// TIA Portal project "python_communication" (V18)

(* hardware
DEVICE "S7-1200 station_1"  S7-1200 Station
   slot 0: "Rack_0"  S7-1200 Rack  Rack  V1.0
   slot 1: "PLC_1"  CPU 1214C DC/DC/Rly  6ES7 214-1HG40-0XB0  V4.6
*)

// ===== PLC "PLC_1"  CPU 1214C DC/DC/Rly =====

VAR_GLOBAL   // PLC tag table "Default tag table"
   "Main_Conveyor_Motor" AT %Q10.0 : Bool;
   "Start_But" AT %I10.0 : Bool;
   "Stop_But" AT %I10.1 : Bool;
   "Start_Mem" AT %M1.0 : Bool;
   "First_Detected_Sensor" AT %I10.2 : Bool;
   "Stop_Mem" AT %M2.0 : Bool;
   "Second_Band_Exit_Sensor" AT %I10.3 : Bool;
   "Second_Band_First_Sensor" AT %I10.4 : Bool;
   "Machine_Sensor" AT %I10.5 : Bool;
   "Move_Z_Mem" AT %M3.0 : Bool;
   "Move_Z" AT %Q10.1 : Bool;
   "Grab_İtem" AT %Q10.2 : Bool;
   "Grab_Mem" AT %M4.0 : Bool;
   "Move_X_Mem" AT %M5.0 : Bool;
   "Move_X" AT %Q10.3 : Bool;
   "Moving_X" AT %I10.6 : Bool;
   "Moving_Z" AT %I10.7 : Bool;
   "Second_Band_Motor" AT %Q10.4 : Bool;
   "Second_Band_Motor_Mem" AT %M6.0 : Bool;
   "Defect_Process_Active" AT %M7.0 : Bool;
   "Corner_Band_Motor" AT %Q10.5 : Bool;
   "Main_Band2_Motor" AT %Q10.6 : Bool;
   "Stack_Light(RED)" AT %Q10.7 : Bool;
   "Stack_Light(GREEN)" AT %Q11.0 : Bool;
   "Stack_Light(YELLOW)" AT %Q11.1 : Bool;
   "Python_Alive" AT %M8.0 : Bool;
END_VAR

DATA_BLOCK "DB_Python"   // DB1
{ S7_Optimized_Access := 'FALSE' }
VERSION : 0.1
   VAR
      Trigger : Bool;
      Part_At_Camera : Bool;
      Heartbeat : Bool;
      DefectCount : Int;
      ConfidenceScore : Real;
   END_VAR
BEGIN
END_DATA_BLOCK

// folder: System blocks/Program resources

DATA_BLOCK "timer5"   // DB2
{ S7_Optimized_Access := 'TRUE' }
AUTHOR : Simatic
FAMILY : IEC
NAME : IEC_TMR
VERSION : 1.0
// stored: InstanceOfName IEC_TIMER
"IEC_TIMER"
BEGIN
END_DATA_BLOCK

DATA_BLOCK "timer1"   // DB3
{ S7_Optimized_Access := 'TRUE' }
AUTHOR : Simatic
FAMILY : IEC
NAME : IEC_TMR
VERSION : 1.0
// stored: InstanceOfName IEC_TIMER
"IEC_TIMER"
BEGIN
END_DATA_BLOCK

DATA_BLOCK "Timer2"   // DB4
{ S7_Optimized_Access := 'TRUE' }
AUTHOR : Simatic
FAMILY : IEC
NAME : IEC_TMR
VERSION : 1.0
// stored: InstanceOfName IEC_TIMER
"IEC_TIMER"
BEGIN
END_DATA_BLOCK

DATA_BLOCK "timer3"   // DB5
{ S7_Optimized_Access := 'TRUE' }
AUTHOR : Simatic
FAMILY : IEC
NAME : IEC_TMR
VERSION : 1.0
// stored: InstanceOfName IEC_TIMER
"IEC_TIMER"
BEGIN
END_DATA_BLOCK

// folder: (top level)

FUNCTION "MHJ-PLC-Lab-Function-S71200" : Void   // FC9000, SCL
{ S7_Optimized_Access := 'TRUE' }
VERSION : 0.1
   VAR_TEMP
      rdTimeReturn : Int;
      outputTime : DTL;
      SyncVal : Byte;
      forVal : Int;
      forVal_2 : Int;
      Value : Byte;
   END_VAR
   VAR CONSTANT
      CompVal : Byte := 16#34;
      Value_01 : Byte := 16#11;
      Value_01_DW : DWord := 16#A165_D992;
      Value_02_DW : DWord := 16#58BE_4401;
   END_VAR
BEGIN

   #Value:=PEEK(area := 16#82,
        dbNumber := 0,
        byteOffset := 511);
   #Value := #Value + 1;

   POKE(area := 16#82,
        dbNumber := 0,
        byteOffset := 511,
        value := #Value);

   POKE(area:=16#81,
        dbNumber:=0,
        byteOffset:=1016,
        value:=#Value_01_DW);
   POKE(area := 16#81,
        dbNumber := 0,
        byteOffset := 1020,
        value := #Value_02_DW);

   POKE(area := 16#81,
        dbNumber := 0,
        byteOffset := 511,
        value := B#16#00);

   FOR #forVal := 0 TO 120 DO
       FOR #forVal_2:=0 TO 10 DO
           #rdTimeReturn:=RD_SYS_T(#outputTime);
           #rdTimeReturn := WR_SYS_T(#outputTime);
           #rdTimeReturn := RD_SYS_T(#outputTime);
           #rdTimeReturn := WR_SYS_T(#outputTime);
       END_FOR;
       #SyncVal:= PEEK(area := 16#81,
                      dbNumber := 0,
                      byteOffset := 511);
       IF #SyncVal = #CompVal THEN
          GOTO M_1;
       END_IF;
   END_FOR;
   RETURN;

   M_1:
   POKE(area := 16#81,
        dbNumber := 0,
        byteOffset := 511,
        value := B#16#0);
END_FUNCTION

ORGANIZATION_BLOCK "Main"   // OB1, LAD, ProgramCycle
TITLE = "Main Program Sweep (Cycle)"
{ S7_Optimized_Access := 'TRUE' }
VERSION : 0.1
   VAR_INPUT
      Initial_Call : Bool;   // Initial call of this OB
      Remanence : Bool;   // =True, if remanent data are available
   END_VAR
   VAR_TEMP   // added for the SCL form of the ladder/FBD networks
      _w1 : Bool;
      _w2 : Bool;
   END_VAR
BEGIN

REGION Network 1: FactoryIO_Communication
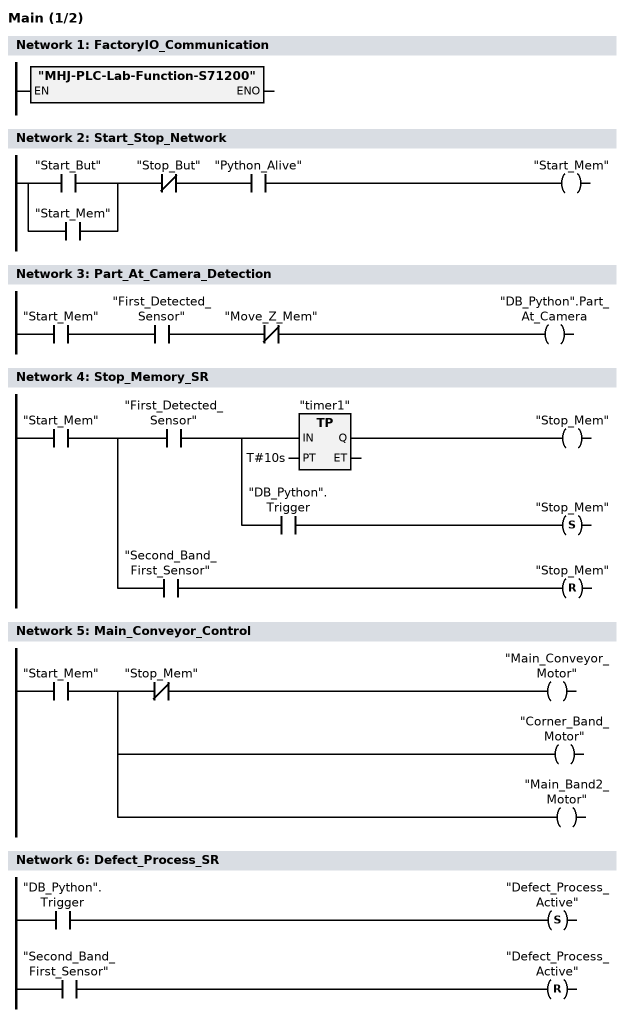
   RUNG wire#powerrail
      "MHJ-PLC-Lab-Function-S71200"()
   END_RUNG
   // the same network as SCL:
   "MHJ-PLC-Lab-Function-S71200"();
END_REGION

REGION Network 2: Start_Stop_Network
   RUNG wire#powerrail
      Contact( "Start_But" )
      wire#w1
      I_Contact( "Stop_But" )
      Contact( "Python_Alive" )
      Coil( "Start_Mem" )
   END_RUNG
   RUNG wire#powerrail
      Contact( "Start_Mem" )
   END_RUNG wire#w1
   // the same network as SCL:
   "Start_Mem" := ("Start_But" OR "Start_Mem") AND NOT "Stop_But" AND "Python_Alive";
END_REGION

REGION Network 3: Part_At_Camera_Detection
   RUNG wire#powerrail
      Contact( "Start_Mem" )
      Contact( "First_Detected_Sensor" )
      I_Contact( "Move_Z_Mem" )
      Coil( "DB_Python".Part_At_Camera )
   END_RUNG
   // the same network as SCL:
   "DB_Python".Part_At_Camera := "Start_Mem" AND "First_Detected_Sensor" AND NOT "Move_Z_Mem";
END_REGION

REGION Network 4: Stop_Memory_SR
   #_w1 := "Start_Mem" AND "First_Detected_Sensor";
   "timer1".TP(IN := #_w1, PT := T#10s);
   "Stop_Mem" := "timer1".Q;
   IF #_w1 AND "DB_Python".Trigger THEN "Stop_Mem" := TRUE; END_IF;
   IF "Start_Mem" AND "Second_Band_First_Sensor" THEN "Stop_Mem" := FALSE; END_IF;
END_REGION

REGION Network 5: Main_Conveyor_Control
   RUNG wire#powerrail
      Contact( "Start_Mem" )
      wire#w1
      I_Contact( "Stop_Mem" )
      Coil( "Main_Conveyor_Motor" )
   END_RUNG
   RUNG wire#w1
      Coil( "Corner_Band_Motor" )
   END_RUNG
   RUNG wire#w1
      Coil( "Main_Band2_Motor" )
   END_RUNG
   // the same network as SCL:
   "Main_Conveyor_Motor" := "Start_Mem" AND NOT "Stop_Mem";
   "Corner_Band_Motor" := "Start_Mem";
   "Main_Band2_Motor" := "Start_Mem";
END_REGION

REGION Network 6: Defect_Process_SR
   RUNG wire#powerrail
      Contact( "DB_Python".Trigger )
      S_Coil( "Defect_Process_Active" )
   END_RUNG
   RUNG wire#powerrail
      Contact( "Second_Band_First_Sensor" )
      R_Coil( "Defect_Process_Active" )
   END_RUNG
   // the same network as SCL:
   IF "DB_Python".Trigger THEN "Defect_Process_Active" := TRUE; END_IF;
   IF "Second_Band_First_Sensor" THEN "Defect_Process_Active" := FALSE; END_IF;
END_REGION

REGION Network 7: Pick_and_Place_State_Machine
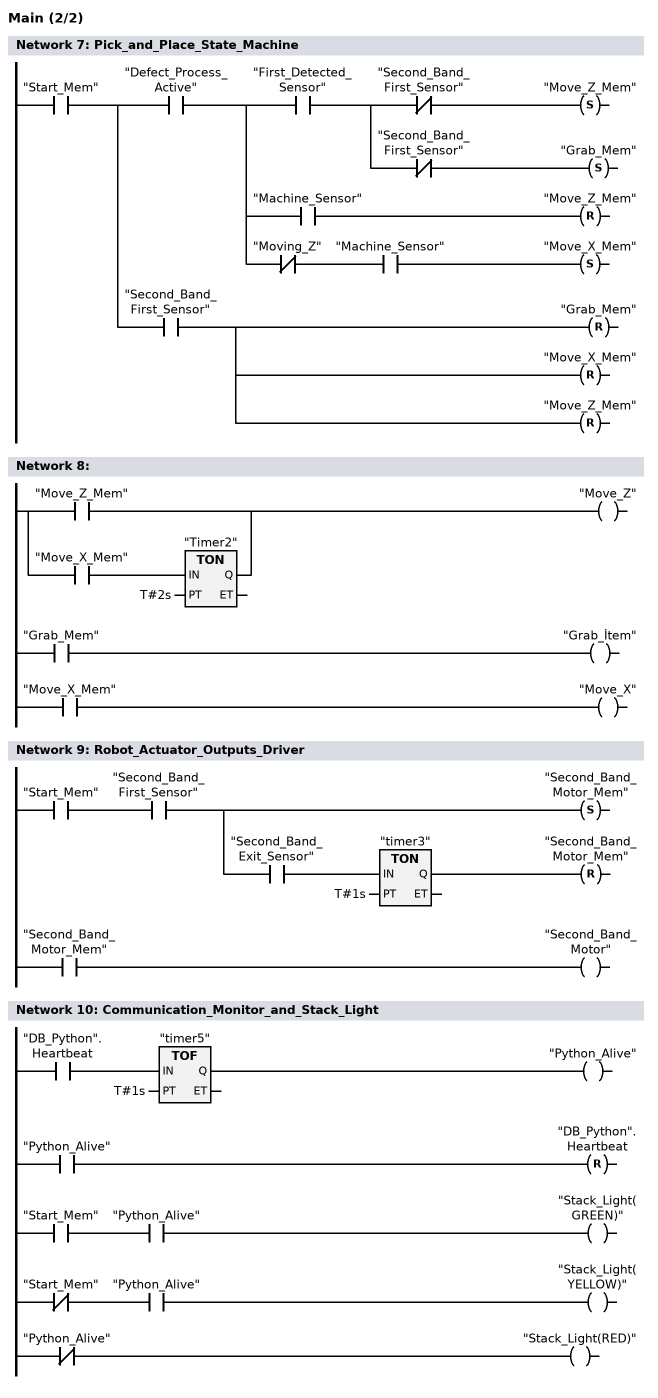
   RUNG wire#powerrail
      Contact( "Start_Mem" )
      wire#w1
      Contact( "Defect_Process_Active" )
      wire#w2
      Contact( "First_Detected_Sensor" )
      wire#w3
      I_Contact( "Second_Band_First_Sensor" )
      S_Coil( "Move_Z_Mem" )
   END_RUNG
   RUNG wire#w3
      I_Contact( "Second_Band_First_Sensor" )
      S_Coil( "Grab_Mem" )
   END_RUNG
   RUNG wire#w2
      Contact( "Machine_Sensor" )
      R_Coil( "Move_Z_Mem" )
   END_RUNG
   RUNG wire#w2
      I_Contact( "Moving_Z" )
      Contact( "Machine_Sensor" )
      S_Coil( "Move_X_Mem" )
   END_RUNG
   RUNG wire#w1
      Contact( "Second_Band_First_Sensor" )
      wire#w4
      R_Coil( "Grab_Mem" )
   END_RUNG
   RUNG wire#w4
      R_Coil( "Move_X_Mem" )
   END_RUNG
   RUNG wire#w4
      R_Coil( "Move_Z_Mem" )
   END_RUNG
   // the same network as SCL:
   #_w1 := "Start_Mem" AND "Defect_Process_Active";
   #_w2 := #_w1 AND "First_Detected_Sensor";
   IF #_w2 AND NOT "Second_Band_First_Sensor" THEN
       "Move_Z_Mem" := TRUE;
       "Grab_Mem" := TRUE;
   END_IF;
   IF #_w1 AND "Machine_Sensor" THEN "Move_Z_Mem" := FALSE; END_IF;
   IF #_w1 AND NOT "Moving_Z" AND "Machine_Sensor" THEN "Move_X_Mem" := TRUE; END_IF;
   IF "Start_Mem" AND "Second_Band_First_Sensor" THEN
       "Grab_Mem" := FALSE;
       "Move_X_Mem" := FALSE;
       "Move_Z_Mem" := FALSE;
   END_IF;
END_REGION

REGION Network 8
   "Timer2".TON(IN := "Move_X_Mem", PT := T#2s);
   "Move_Z" := "Move_Z_Mem" OR "Timer2".Q;
   "Grab_İtem" := "Grab_Mem";
   "Move_X" := "Move_X_Mem";
END_REGION

REGION Network 9: Robot_Actuator_Outputs_Driver
   #_w1 := "Start_Mem" AND "Second_Band_First_Sensor";
   IF #_w1 THEN "Second_Band_Motor_Mem" := TRUE; END_IF;
   "timer3".TON(IN := #_w1 AND "Second_Band_Exit_Sensor", PT := T#1s);
   IF "timer3".Q THEN "Second_Band_Motor_Mem" := FALSE; END_IF;
   "Second_Band_Motor" := "Second_Band_Motor_Mem";
END_REGION

REGION Network 10: Communication_Monitor_and_Stack_Light
   "timer5".TOF(IN := "DB_Python".Heartbeat, PT := T#1s);
   "Python_Alive" := "timer5".Q;
   IF "Python_Alive" THEN "DB_Python".Heartbeat := FALSE; END_IF;
   "Stack_Light(GREEN)" := "Start_Mem" AND "Python_Alive";
   "Stack_Light(YELLOW)" := NOT "Start_Mem" AND "Python_Alive";
   "Stack_Light(RED)" := NOT "Python_Alive";
END_REGION
END_ORGANIZATION_BLOCK